(* IEC 61131-3 sources: llm-plc-st-eval/data/definitivo/qwen2.5-coder_14b/I7/few_shot, 3 files *)

(* ---- ejec_1.st ---- *)
FUNCTION_BLOCK FB_Duplex
VAR_INPUT
    demanda : BOOL; (* Demanda de arranque *)
    falla1 : BOOL; (* Falla de la bomba 1 *)
    falla2 : BOOL; (* Falla de la bomba 2 *)
END_VAR
VAR_OUTPUT
    bomba1 : BOOL; (* Bomba principal *)
    bomba2 : BOOL; (* Bomba secundaria *)
    almFalla : BOOL; (* Alarma de falla de la bomba principal *)
END_VAR
VAR
    estado : INT := 0; (* Estado del sistema *)
    cambio : BOOL := FALSE; (* Bandera de cambio de estado *)
END_VAR

(* Estado 0: Espera inicial *)
IF demanda THEN
    estado := 1;
    cambio := TRUE;
END_IF

(* Estado 1: Bomba 1 principal *)
IF estado = 1 THEN
    IF NOT falla1 THEN
        bomba1 := TRUE;
        bomba2 := FALSE;
        almFalla := FALSE;
    ELSE
        IF NOT falla2 THEN
            bomba1 := FALSE;
            bomba2 := TRUE;
            almFalla := TRUE;
        ELSE
            bomba1 := FALSE;
            bomba2 := FALSE;
            almFalla := TRUE;
        END_IF
    END_IF
END_IF

(* Estado 2: Bomba 2 principal *)
IF estado = 2 THEN
    IF NOT falla2 THEN
        bomba1 := FALSE;
        bomba2 := TRUE;
        almFalla := FALSE;
    ELSE
        IF NOT falla1 THEN
            bomba1 := TRUE;
            bomba2 := FALSE;
            almFalla := TRUE;
        ELSE
            bomba1 := FALSE;
            bomba2 := FALSE;
            almFalla := TRUE;
        END_IF
    END_IF
END_IF

(* Cambio de estado en nueva demanda *)
IF demanda AND cambio THEN
    IF estado = 1 THEN
        estado := 2;
    ELSE
        estado := 1;
    END_IF
    cambio := FALSE;
END_IF

(* Detener bombas al quitar demanda *)
IF NOT demanda THEN
    bomba1 := FALSE;
    bomba2 := FALSE;
    cambio := TRUE;
END_IF

END_FUNCTION_BLOCK

(* ---- ejec_2.st ---- *)
FUNCTION_BLOCK FB_Duplex
VAR_INPUT
    demanda : BOOL; (* Demanda de arranque *)
    falla1 : BOOL; (* Falla de la bomba 1 *)
    falla2 : BOOL; (* Falla de la bomba 2 *)
END_VAR
VAR_OUTPUT
    bomba1 : BOOL; (* Bomba principal *)
    bomba2 : BOOL; (* Bomba de respaldo *)
    almFalla : BOOL; (* Alarma de falla de la bomba principal *)
END_VAR
VAR
    estado : INT := 0; (* Estado del sistema: 0 - detenido, 1 - bomba1 principal, 2 - bomba2 principal *)
    demandaAnterior : BOOL := FALSE; (* Estado anterior de la demanda *)
END_VAR

(* Cambio de estado en la transición de FALSE a TRUE de demanda *)
IF demanda AND NOT demandaAnterior THEN
    estado := (estado + 1) MOD 3;
END_IF

(* Asignación de bombas según el estado *)
CASE estado OF
    0: (* Detenido *)
        bomba1 := FALSE;
        bomba2 := FALSE;
    1: (* Bomba1 principal *)
        bomba1 := NOT falla1;
        bomba2 := falla1 AND NOT falla2;
    2: (* Bomba2 principal *)
        bomba1 := falla2 AND NOT falla1;
        bomba2 := NOT falla2;
END_CASE

(* Alarma de falla de la bomba principal *)
almFalla := (estado = 1 AND falla1) OR (estado = 2 AND falla2);

(* Actualización del estado anterior de la demanda *)
demandaAnterior := demanda;
END_FUNCTION_BLOCK

(* ---- ejec_3.st ---- *)
FUNCTION_BLOCK FB_Duplex
VAR_INPUT
    demanda : BOOL; (* Demanda de arranque *)
    falla1 : BOOL; (* Falla de la bomba 1 *)
    falla2 : BOOL; (* Falla de la bomba 2 *)
END_VAR
VAR_OUTPUT
    bomba1 : BOOL; (* Bomba principal *)
    bomba2 : BOOL; (* Bomba de respaldo *)
    almFalla : BOOL; (* Alarma de falla de la bomba principal *)
END_VAR
VAR
    estado : INT := 0; (* Estado actual: 0 = detenido, 1 = bomba1 principal, 2 = bomba2 principal *)
    demandaAnterior : BOOL := FALSE; (* Estado anterior de la demanda *)
END_VAR

(* Control de la alternancia de bombas y manejo de fallas *)
IF demanda THEN
    IF NOT demandaAnterior THEN
        (* Transición de FALSE a TRUE en demanda *)
        estado := (estado + 1) MOD 3;
        IF estado = 0 THEN
            estado := 1; (* Asegura que la primera demanda arranque bomba1 *)
        END_IF
    END_IF

    CASE estado OF
        1:
            IF falla1 THEN
                bomba1 := FALSE;
                bomba2 := NOT falla2;
                almFalla := NOT falla2;
            ELSE
                bomba1 := TRUE;
                bomba2 := FALSE;
                almFalla := FALSE;
            END_IF
        2:
            IF falla2 THEN
                bomba2 := FALSE;
                bomba1 := NOT falla1;
                almFalla := NOT falla1;
            ELSE
                bomba2 := TRUE;
                bomba1 := FALSE;
                almFalla := FALSE;
            END_IF
    END_CASE
ELSE
    bomba1 := FALSE;
    bomba2 := FALSE;
    almFalla := FALSE;
END_IF

(* Actualización del estado anterior de la demanda *)
demandaAnterior := demanda;
END_FUNCTION_BLOCK
